# EPICS substitutions: iocs/motor/esp300-ioc/db/ESP300.substitutions
# C's iocNewport ESP300.substitutions, P from st.cmd.
file "$(MOTOR)/db/motor.db"
{
pattern
{N,   M,        DTYP,      C,  S,  DESC,          EGU,  DIR,  VELO,  VBAS,  ACCL,  BDST,  BVEL,  BACC,  MRES,  PREC,  DHLM,  DLLM,  INIT}
{21,  "m$(N)",  "ESP300",  0,  0,  "motor $(N)",  mm,   Pos,  1,     .1,    .2,    0,     1,     .2,    5e-5,  5,     100,   -100,  ""}
{22,  "m$(N)",  "ESP300",  0,  1,  "motor $(N)",  mm,   Pos,  1,     .1,    .2,    0,     1,     .2,    5e-5,  5,     100,   -100,  ""}
{23,  "m$(N)",  "ESP300",  0,  2,  "motor $(N)",  mm,   Pos,  1,     .1,    .2,    0,     1,     .2,    5e-5,  5,     100,   -100,  ""}
}
